Fanuc KAREL source: kc00038.KL

-- PROVISIONAL review KL for V940-1; original PC SHA256 7967f3562545c9e7e5250c176f94237fd4879baaed34b7a0e26c8aeff7e77117
-- Incomplete behavior may be omitted. Consult companion uncertainty JSON. Do not deploy.
PROGRAM KC00038
%NOLOCKGROUP
BEGIN
  -- V9_ZERO_TABLE_METADATA_HINT layout=0001; no indexed target words; source/name/runtime held
  -- UNRESOLVED_PC offsets 5-32; opcodes 27,22,1C,22,22,76
  -- UNRESOLVED_PC offsets 37-41; opcodes 7F
END KC00038
